// Generated by voz_llm_plc_agent
// Target: Siemens TIA Portal V18 - SCL external source
// Review and compile before any download to physical hardware.

FUNCTION_BLOCK "PLC_PRG"
{ S7_Optimized_Access := 'TRUE' }
VERSION : 0.1
VAR_INPUT
   I_Start : Bool := FALSE;
   I_Reset : Bool := FALSE;
   I_Emergency : Bool := FALSE;
END_VAR
VAR_OUTPUT
   Q_Motor_Enable : Bool := FALSE;
   Q_Cycle_Complete : Bool := FALSE;
END_VAR
VAR
   M_CycleStep : Bool;
   T_Cycle {InstructionName := 'TON_TIME'; LibVersion := '1.0'} : TON_TIME;
END_VAR
BEGIN
(* Ciclo automatico temporizado: 0 = inicial, 1 = en ejecucion, 2 = finalizado (hasta Reset) *)
IF #I_Emergency OR #I_Reset THEN
    #M_CycleStep := 0;
ELSIF #M_CycleStep = 0 AND #I_Start THEN
    #M_CycleStep := 1;
END_IF;

#T_Cycle(IN := #M_CycleStep = 1, PT := T#3s);
IF #M_CycleStep = 1 AND #T_Cycle.Q THEN
    #M_CycleStep := 2;
END_IF;

#Q_Motor_Enable := #M_CycleStep = 1 AND NOT #I_Emergency;
#Q_Cycle_Complete := #M_CycleStep = 2;
(* Bloqueo: #I_Emergency fuerza a FALSE #Q_Motor_Enable de inmediato *)
IF #I_Emergency THEN
    #Q_Motor_Enable := FALSE;
END_IF;
END_FUNCTION_BLOCK

DATA_BLOCK "DB_PLC_PRG"
{ S7_Optimized_Access := 'TRUE' }
VERSION : 0.1
NON_RETAIN
"PLC_PRG"
BEGIN
END_DATA_BLOCK

ORGANIZATION_BLOCK "Main"
{ S7_Optimized_Access := 'TRUE' }
VERSION : 0.1
BEGIN
   "DB_PLC_PRG"(
      I_Start := "I_Start",
      I_Reset := "I_Reset",
      I_Emergency := "I_Emergency",
      Q_Motor_Enable => "Q_Motor_Enable",
      Q_Cycle_Complete => "Q_Cycle_Complete"
   );
END_ORGANIZATION_BLOCK
